(* IEC 61131-3 sources: llm-plc-st-eval/data/processed_definitivo/claude-sonnet-4-6/A4/zero_shot, 3 files *)

(* ---- ejec_1.st ---- *)
FUNCTION_BLOCK FB_Rampa
VAR_INPUT
    SPvel     : REAL; (* Consigna de velocidad [%] *)
    paroRapido: BOOL; (* Paro rápido activo *)
    ciclo     : TIME; (* Período de ejecución del bloque *)
END_VAR

VAR_OUTPUT
    CVvel : REAL; (* Salida de velocidad con rampa [%] *)
END_VAR

VAR
    rSegundos   : REAL; (* Período en segundos *)
    rMaxSubida  : REAL; (* Incremento máximo por ciclo al subir *)
    rMaxBajada  : REAL; (* Decremento máximo por ciclo al bajar *)
    rMaxParada  : REAL; (* Decremento máximo por ciclo en paro rápido *)
    rError      : REAL; (* Diferencia entre SP y CV *)
END_VAR

(* ── Constantes de pendiente [puntos porcentuales / segundo] ── *)
CONST
    PENDIENTE_SUBIDA : REAL := 10.0;
    PENDIENTE_BAJADA : REAL := 20.0;
    PENDIENTE_PARO   : REAL := 40.0;
END_CONST

(* ── Conversión del período de ciclo a segundos ── *)
rSegundos := TIME_TO_REAL(ciclo) / 1000.0;

(* ── Incrementos máximos permitidos en este ciclo ── *)
rMaxSubida := PENDIENTE_SUBIDA * rSegundos;
rMaxBajada := PENDIENTE_BAJADA * rSegundos;
rMaxParada := PENDIENTE_PARO  * rSegundos;

IF paroRapido THEN
    (* ── Paro rápido: descender hacia 0.0 ignorando SPvel ── *)
    IF CVvel > 0.0 THEN
        CVvel := CVvel - rMaxParada;
        IF CVvel < 0.0 THEN
            CVvel := 0.0; (* Sin sobrepaso por debajo de 0 *)
        END_IF;
    ELSIF CVvel < 0.0 THEN
        (* Si por alguna razón CV fuera negativo, llevarlo a 0 *)
        CVvel := CVvel + rMaxParada;
        IF CVvel > 0.0 THEN
            CVvel := 0.0;
        END_IF;
    END_IF;
    (* Mientras paroRapido siga activo y CV = 0, permanece en 0 *)
ELSE
    (* ── Seguimiento normal de la consigna con rampa ── *)
    rError := SPvel - CVvel;

    IF rError > 0.0 THEN
        (* Subida: limitar el incremento a rMaxSubida *)
        CVvel := CVvel + rMaxSubida;
        IF CVvel > SPvel THEN
            CVvel := SPvel; (* Sin sobrepaso por arriba *)
        END_IF;

    ELSIF rError < 0.0 THEN
        (* Bajada: limitar el decremento a rMaxBajada *)
        CVvel := CVvel - rMaxBajada;
        IF CVvel < SPvel THEN
            CVvel := SPvel; (* Sin sobrepaso por abajo *)
        END_IF;

    (* Si rError = 0.0, CVvel ya es igual a SPvel; no se hace nada *)
    END_IF;
END_IF;

END_FUNCTION_BLOCK

(* ---- ejec_2.st ---- *)
FUNCTION_BLOCK FB_Rampa
VAR_INPUT
    SPvel     : REAL;   (* Consigna de velocidad [%] *)
    paroRapido: BOOL;   (* Paro rápido activo *)
    ciclo     : TIME;   (* Período de ejecución del bloque *)
END_VAR

VAR_OUTPUT
    CVvel : REAL;       (* Salida de velocidad con rampa [%] *)
END_VAR

VAR
    rSegundos  : REAL;  (* Período de ciclo convertido a segundos *)
    rMaxSubida : REAL;  (* Incremento máximo permitido en un ciclo *)
    rMaxBajada : REAL;  (* Decremento máximo permitido en un ciclo *)
    rError     : REAL;  (* Diferencia entre consigna y salida actual *)
END_VAR

(* ── Constantes de pendiente [puntos porcentuales / segundo] ── *)
VAR CONSTANT
    PENDIENTE_SUBIDA    : REAL := 10.0;
    PENDIENTE_BAJADA    : REAL := 20.0;
    PENDIENTE_PARO_RAP  : REAL := 40.0;
END_VAR

(* ── Conversión del período de ciclo a segundos ── *)
rSegundos := TIME_TO_REAL(ciclo) / 1000.0;

IF paroRapido THEN
    (* ── Modo paro rápido: descender hacia 0.0 con pendiente rápida ── *)
    rMaxBajada := PENDIENTE_PARO_RAP * rSegundos;

    IF CVvel > 0.0 THEN
        CVvel := CVvel - rMaxBajada;
        (* Evitar sobrepaso por debajo de 0.0 *)
        IF CVvel < 0.0 THEN
            CVvel := 0.0;
        END_IF;
    ELSE
        (* Mantener en 0.0 mientras paroRapido siga activo *)
        CVvel := 0.0;
    END_IF;

ELSE
    (* ── Modo normal: seguir SPvel con pendientes limitadas ── *)
    rMaxSubida := PENDIENTE_SUBIDA * rSegundos;
    rMaxBajada := PENDIENTE_BAJADA * rSegundos;

    rError := SPvel - CVvel;

    IF rError > 0.0 THEN
        (* Consigna mayor que salida: subir con pendiente limitada *)
        IF rError > rMaxSubida THEN
            CVvel := CVvel + rMaxSubida;
        ELSE
            (* El paso restante es menor que el máximo: llegar exactamente *)
            CVvel := SPvel;
        END_IF;

    ELSIF rError < 0.0 THEN
        (* Consigna menor que salida: bajar con pendiente limitada *)
        IF (-rError) > rMaxBajada THEN
            CVvel := CVvel - rMaxBajada;
        ELSE
            CVvel := SPvel;
        END_IF;

    (* Si rError = 0.0, CVvel ya es igual a SPvel; no se hace nada *)
    END_IF;

END_IF;

END_FUNCTION_BLOCK

(* ---- ejec_3.st ---- *)
FUNCTION_BLOCK FB_Rampa
VAR_INPUT
    SPvel     : REAL;   (* Consigna de velocidad [%] *)
    paroRapido: BOOL;   (* Paro rápido activo *)
    ciclo     : TIME;   (* Período de ejecución del bloque *)
END_VAR

VAR_OUTPUT
    CVvel : REAL;       (* Salida de velocidad con rampa [%] *)
END_VAR

VAR
    rPendiente  : REAL; (* Pendiente aplicada en este ciclo [puntos/%] *)
    rDelta      : REAL; (* Incremento/decremento máximo en este ciclo *)
    rSegundos   : REAL; (* Período de ciclo convertido a segundos *)
    rObjetivo   : REAL; (* Valor objetivo en este ciclo *)
END_VAR

(* ── Constantes de rampa [puntos porcentuales / segundo] ── *)
VAR CONSTANT
    C_RAMPA_SUBIDA  : REAL := 10.0;  (* Máx. subida  *)
    C_RAMPA_BAJADA  : REAL := 20.0;  (* Máx. bajada  *)
    C_RAMPA_PARO    : REAL := 40.0;  (* Paro rápido  *)
END_VAR

(* ── Conversión del período a segundos ── *)
rSegundos := TIME_TO_REAL(ciclo) / 1000.0;

IF paroRapido THEN
    (* ── Modo paro rápido: descender hacia 0.0 con rampa de 40 %/s ── *)
    rObjetivo := 0.0;

    IF CVvel > 0.0 THEN
        (* Calcular decremento máximo permitido en este ciclo *)
        rDelta := C_RAMPA_PARO * rSegundos;
        CVvel  := CVvel - rDelta;

        (* Evitar sobrepasar el objetivo (0.0) por debajo *)
        IF CVvel < 0.0 THEN
            CVvel := 0.0;
        END_IF;

    ELSIF CVvel < 0.0 THEN
        (* Si por alguna razón CVvel es negativo, subir hacia 0.0 *)
        rDelta := C_RAMPA_PARO * rSegundos;
        CVvel  := CVvel + rDelta;

        IF CVvel > 0.0 THEN
            CVvel := 0.0;
        END_IF;

    END_IF;
    (* CVvel = 0.0 exacto: no se modifica *)

ELSE
    (* ── Modo normal: seguir SPvel con rampa de subida/bajada ── *)
    rObjetivo := SPvel;

    IF CVvel < rObjetivo THEN
        (* Subida: pendiente limitada a C_RAMPA_SUBIDA *)
        rDelta := C_RAMPA_SUBIDA * rSegundos;
        CVvel  := CVvel + rDelta;

        (* Evitar sobrepasar el objetivo por arriba *)
        IF CVvel > rObjetivo THEN
            CVvel := rObjetivo;
        END_IF;

    ELSIF CVvel > rObjetivo THEN
        (* Bajada: pendiente limitada a C_RAMPA_BAJADA *)
        rDelta := C_RAMPA_BAJADA * rSegundos;
        CVvel  := CVvel - rDelta;

        (* Evitar sobrepasar el objetivo por abajo *)
        IF CVvel < rObjetivo THEN
            CVvel := rObjetivo;
        END_IF;

    END_IF;
    (* CVvel = rObjetivo exacto: no se modifica *)

END_IF;
